{attribute 'qualified_only'}
VAR_GLOBAL PERSISTENT
	platform : PlatformKind := PlatformKind.SIMULATION;
	// Hjulradien ligger i NC-skaleringen av aksene, som går i meter langs hjulbanen.
	trackWidthInM : LREAL := 0.40;
	maxWheelSpeedInMPerS : LREAL := 0.6;
END_VAR

(* stored: Version 1.1.0.1, ProductVersion 3.1.4026.12
   GVL Parameters: Id {1597954a-e0f8-5851-b29a-c1b34e85d36f} *)
